FUNCTION_BLOCK "FB1062_HorDrillAutoStep"   // FB1062, SCL
{ S7_Optimized_Access := 'TRUE' }
// ============================================================
//  Block: FB1062_HorDrillAutoStep
//  ============================================================
//  编号：FB1062
//  原始语言：LAD（规则翻译为 SCL）
//  含义：Added Visual Chiseling Modeby WXY, 20220727
   VAR
      Aux : Struct   // 静态变量
         StartDrill : Bool;   // 静态变量
         DrillDepthMid : DInt;   // 打孔深度中间变量
         DrillDepthMax : Real;   // 静态变量
         DrillDepthMin : Real;   // 静态变量
         ScrLen_Mid : DInt;   // 批头长度中间变量
         OffSetYMid : DInt;   // 静态变量
         OffSetZMid : DInt;   // 静态变量
         go_X : Real;   // 机器人当前X位置
         go_Z : Real;   // 机器人当前Z位置
         MidPos_X : DInt;   // 静态变量
         MidPos_Z : DInt;   // 静态变量
         RobotSpeed : DInt;   // 机器人速度写入
         PressureMid : Real;   // 力中间变量
         HDrillOutTime : IEC_TIMER;   // 水平钻孔超时
         HStartTime : IEC_TIMER;   // 水平钻孔超时
      END_STRUCT;
      EdgeDetc : Struct   // 静态变量
         Pulse : Array[0..15] of Bool;   // 静态变量
      END_STRUCT;
      HorDrillStep : Struct   // 水平钻孔
         Busy : Bool;   // 静态变量
         StartCmd : Bool;   // 静态变量
         OKToStart : Bool;   // 静态变量
         TaskDone : Bool;   // 静态变量
         StepStart : Bool;   // 静态变量
         StepEnd : Bool;   // 静态变量
         ErrEnd : Bool;   // 静态变量
         ByPass : Bool;   // 静态变量
         TaskIO : Bool;   // 静态变量
         TaskNIO : Bool;   // 静态变量
         S1 : Bool;   // 静态变量
         S2 : Bool;   // 静态变量
         S3 : Bool;   // 静态变量
         S4 : Bool;   // 静态变量
         S5 : Bool;   // 静态变量
         S6 : Bool;   // 静态变量
         S7 : Bool;   // 静态变量
         S8 : Bool;   // 静态变量
         S9 : Bool;   // 静态变量
         S10 : Bool;   // 静态变量
         S11 : Bool;   // 静态变量
         S12 : Bool;   // 静态变量
         S13 : Bool;   // 静态变量
         S14 : Bool;   // 静态变量
         S15 : Bool;   // 静态变量
         S16 : Bool;   // 静态变量
         S17 : Bool;   // 静态变量
         S18 : Bool;   // 静态变量
         S19 : Bool;   // 静态变量
         S20 : Bool;   // 静态变量
         S21 : Bool;   // 静态变量
         S22 : Bool;   // 静态变量
         S23 : Bool;   // 静态变量
         S24 : Bool;   // 静态变量
         S25 : Bool;   // 静态变量
         S26 : Bool;   // 静态变量
         S27 : Bool;   // 静态变量
         S28 : Bool;   // 静态变量
         S29 : Bool;   // 静态变量
         S30 : Bool;   // 静态变量
         S31 : Bool;   // 静态变量
         S32 : Bool;   // 静态变量
         S33 : Bool;   // 静态变量
         S34 : Bool;   // 静态变量
         S35 : Bool;   // 静态变量
         S36 : Bool;   // 静态变量
         S37 : Bool;   // 静态变量
         S38 : Bool;   // 静态变量
         S39 : Bool;   // 静态变量
         S40 : Bool;   // 静态变量
         S41 : Bool;   // 静态变量
         S42 : Bool;   // 静态变量
         S43 : Bool;   // 静态变量
         S44 : Bool;   // 静态变量
         S45 : Bool;   // 静态变量
         S46 : Bool;   // 静态变量
         S47 : Bool;   // 静态变量
         S48 : Bool;   // 静态变量
         S49 : Bool;   // 静态变量
         S50 : Bool;   // 静态变量
         S51 : Bool;   // 静态变量
         S52 : Bool;   // 静态变量
         S53 : Bool;   // 静态变量
         S54 : Bool;   // 静态变量
         S55 : Bool;   // 静态变量
         S56 : Bool;   // 静态变量
         S57 : Bool;   // 静态变量
         S58 : Bool;   // 静态变量
         S59 : Bool;   // 静态变量
         S60 : Bool;   // 静态变量
         S61 : Bool;   // 静态变量
         S62 : Bool;   // 静态变量
         S63 : Bool;   // 静态变量
         S64 : Bool;   // 静态变量
         S65 : Bool;   // 静态变量
         S66 : Bool;   // 静态变量
         S67 : Bool;   // 静态变量
         StopDrill_Ack : Bool;   // 静态变量
         GougeStopDrill_Ack : Bool;   // 斜打结束请求
         StopDrill_End : Bool;   // 静态变量
         GougeStopDrill_End : Bool;   // 斜打异常结束请求
         InitForcePulse : Bool;   // 静态变量
      END_STRUCT;
      VisualOffsetMid : Struct   // 静态变量
         X : DInt;   // 静态变量
         Y : DInt;   // 静态变量
         Z : DInt;   // 静态变量
         "A" : DInt;   // 静态变量
         "B" : DInt;   // 静态变量
         C : DInt;   // 静态变量
         A0 : Real;   // 静态变量
         B0 : Real;   // 静态变量
         C0 : Real;   // 静态变量
      END_STRUCT;
      PT : Time;   // 静态变量
      ET : Time;   // 静态变量
      IN : Bool;   // 静态变量
      Q : Bool;   // 水平钻孔超时
   END_VAR
   VAR_TEMP
      StepPls : Bool;   // 临时变量
      HorPosMod : Int;   // 临时变量
   END_VAR
BEGIN

   // ---------- 网络 1 ----------
   // 标题：本工位必须要做(可能条件暂时不满足)
   // 含义：将 (("DB720_KuKa_MainCtrl".Ctrl_Out.RobotAction = 0) AND "DB720_KuKa_MainCtrl".Aux.ToolAtPos) AND NOT ("DB1148_PromptBeeper".Public.RobotNotReady) 赋给 #HorDrillStep.OKToStart
   #HorDrillStep.OKToStart := (("DB720_KuKa_MainCtrl".Ctrl_Out.RobotAction = 0) AND "DB720_KuKa_MainCtrl".Aux.ToolAtPos) AND NOT ("DB1148_PromptBeeper".Public.RobotNotReady);
   // 含义：条件 (("ManMode_M" AND "DB1900_Communication_PC".Recv.RobotDrillTPPB) AND ("DB1900_Communication_PC".Recv.ChooseProgNo = 1)) 成立时，将 TRUE 传送到 #HorDrillStep.StartCmd
   IF (("ManMode_M" AND "DB1900_Communication_PC".Recv.RobotDrillTPPB) AND ("DB1900_Communication_PC".Recv.ChooseProgNo = 1)) THEN
       #HorDrillStep.StartCmd := TRUE;
   END_IF;
   // 含义：将 "DB1900_Communication_PC".Para.DrillDepth; (* Convert → DInt *) END_IF 赋给 IF "DB1060_AutoStep".DownDrillAutoStep.DownDrillStep.StepStart THEN #Aux.DrillDepthMid
   IF "DB1060_AutoStep".DownDrillAutoStep.DownDrillStep.StepStart THEN
       #Aux.DrillDepthMid := "DB1900_Communication_PC".Para.DrillDepth; (* Convert → DInt *)
   END_IF;
   // 含义：将 SWAP(#Aux.DrillDepthMid) 赋给 "DB720_KuKa_MainCtrl".CmdOut.gi_Depth
   "DB720_KuKa_MainCtrl".CmdOut.gi_Depth := SWAP(#Aux.DrillDepthMid);
   // 含义：条件 #HorDrillStep.StepStart AND "DB1900_Communication_PC".Para.ProduceMode3 成立时，将 ("DB1900_Communication_PC".Para.DrillDepth + 0.0) 传送到 #Aux.DrillDepthMid
   IF #HorDrillStep.StepStart AND "DB1900_Communication_PC".Para.ProduceMode3 THEN
       #Aux.DrillDepthMid := ("DB1900_Communication_PC".Para.DrillDepth + 0.0);
   END_IF;
   // 含义：将 SWAP(#Aux.DrillDepthMid) 赋给 "DB720_KuKa_MainCtrl".CmdOut.gi_Depth
   "DB720_KuKa_MainCtrl".CmdOut.gi_Depth := SWAP(#Aux.DrillDepthMid);
   // 含义：条件 #HorDrillStep.StepStart AND "DB1900_Communication_PC".Para.ProduceMode3 成立时，将 "DB1910_DrillData".AUX.LayerNo 传送到 "DB720_KuKa_MainCtrl".CmdOut.gi_LayerNum
   IF #HorDrillStep.StepStart AND "DB1900_Communication_PC".Para.ProduceMode3 THEN
       "DB720_KuKa_MainCtrl".CmdOut.gi_LayerNum := "DB1910_DrillData".AUX.LayerNo;
   END_IF;
   // 含义：条件 #HorDrillStep.StepStart AND NOT ("DB1900_Communication_PC".Para.ProduceMode3) 成立时，将 ("DB1900_Communication_PC".Para.DrillDepth + 5.0) 传送到 #Aux.DrillDepthMid
   IF #HorDrillStep.StepStart AND NOT ("DB1900_Communication_PC".Para.ProduceMode3) THEN
       #Aux.DrillDepthMid := ("DB1900_Communication_PC".Para.DrillDepth + 5.0);
   END_IF;
   // 含义：将 SWAP(#Aux.DrillDepthMid) 赋给 "DB720_KuKa_MainCtrl".CmdOut.gi_Depth
   "DB720_KuKa_MainCtrl".CmdOut.gi_Depth := SWAP(#Aux.DrillDepthMid);
   // 含义：将 "DB1900_Communication_PC".Para.ScrLen; (* Convert → DInt *) 赋给 #Aux.ScrLen_Mid
   #Aux.ScrLen_Mid := "DB1900_Communication_PC".Para.ScrLen; (* Convert → DInt *)
   // 含义：将 SWAP(#Aux.ScrLen_Mid) 赋给 "DB720_KuKa_MainCtrl".CmdOut.gi_ScrewLength
   "DB720_KuKa_MainCtrl".CmdOut.gi_ScrewLength := SWAP(#Aux.ScrLen_Mid);

   // ---------- 网络 2 ----------
   // 标题：****************************机器人坐标数据传递 深度计算*********************************
   // 注释：Added Visual Chiseling Modeby WXY, 20220727
   // 含义：将 SWAP("DB720_KuKa_MainCtrl".StatusIn.go_X) 赋给 #Aux.MidPos_X
   #Aux.MidPos_X := SWAP("DB720_KuKa_MainCtrl".StatusIn.go_X);
   // 含义：将 #Aux.MidPos_X; (* Convert → Real *) 赋给 #Aux.go_X
   #Aux.go_X := #Aux.MidPos_X; (* Convert → Real *)
   // 含义：将 (#Aux.go_X / 1000.0) 赋给 "DB720_KuKa_MainCtrl".Aux.go_X
   "DB720_KuKa_MainCtrl".Aux.go_X := (#Aux.go_X / 1000.0);
   // 含义：将 SWAP("DB720_KuKa_MainCtrl".StatusIn.go_Z) 赋给 #Aux.MidPos_Z
   #Aux.MidPos_Z := SWAP("DB720_KuKa_MainCtrl".StatusIn.go_Z);
   // 含义：将 #Aux.MidPos_Z; (* Convert → Real *) 赋给 #Aux.go_Z
   #Aux.go_Z := #Aux.MidPos_Z; (* Convert → Real *)
   // 含义：将 (#Aux.go_Z / 1000.0) 赋给 "DB720_KuKa_MainCtrl".Aux.go_Z
   "DB720_KuKa_MainCtrl".Aux.go_Z := (#Aux.go_Z / 1000.0);
   // 含义：条件 (((#HorDrillStep.S12 AND "DB720_KuKa_MainCtrl".StatusIn.do_DrillReady_Act) AND "DB720_KuKa_MainCtrl".StatusIn.do_HorDril_Pos) OR (((((#HorDrillStep.S12 AND "DB720_KuKa_MainCtrl".StatusIn.do_DrillReady_Act) AND "DB2500 Visual Chiseling".VisualChiselingMode) AND "DB720_KuKa_MainCtrl".StatusIn.do_Gouge_Pos) AND ("DB1900_Communication_PC".Recv.Current_2 > "DB1900_Communication_PC".Para.CurrentMinLimit))) OR ((#HorDrillStep.S12 AND NOT (#HorDrillStep.S22)) AND #Aux.StartDrill)) AND NOT (#Aux.StartDrill) 成立时，将 "DB720_KuKa_MainCtrl".Aux.go_X 传送到 "DB720_KuKa_MainCtrl".Aux.XZeroPos
   IF (((#HorDrillStep.S12 AND "DB720_KuKa_MainCtrl".StatusIn.do_DrillReady_Act) AND "DB720_KuKa_MainCtrl".StatusIn.do_HorDril_Pos) OR (((((#HorDrillStep.S12 AND "DB720_KuKa_MainCtrl".StatusIn.do_DrillReady_Act) AND "DB2500 Visual Chiseling".VisualChiselingMode) AND "DB720_KuKa_MainCtrl".StatusIn.do_Gouge_Pos) AND ("DB1900_Communication_PC".Recv.Current_2 > "DB1900_Communication_PC".Para.CurrentMinLimit))) OR ((#HorDrillStep.S12 AND NOT (#HorDrillStep.S22)) AND #Aux.StartDrill)) AND NOT (#Aux.StartDrill) THEN
       "DB720_KuKa_MainCtrl".Aux.XZeroPos := "DB720_KuKa_MainCtrl".Aux.go_X;
   END_IF;
   // 含义：条件 ((#HorDrillStep.S12 AND "DB720_KuKa_MainCtrl".StatusIn.do_DrillReady_Act) AND "DB720_KuKa_MainCtrl".StatusIn.do_HorDril_Pos) OR (((((#HorDrillStep.S12 AND "DB720_KuKa_MainCtrl".StatusIn.do_DrillReady_Act) AND "DB2500 Visual Chiseling".VisualChiselingMode) AND "DB720_KuKa_MainCtrl".StatusIn.do_Gouge_Pos) AND ("DB1900_Communication_PC".Recv.Current_2 > "DB1900_Communication_PC".Para.CurrentMinLimit))) OR ((#HorDrillStep.S12 AND NOT (#HorDrillStep.S22)) AND #Aux.StartDrill) 成立时，将 ("DB720_KuKa_MainCtrl".Aux.go_X - "DB720_KuKa_MainCtrl".Aux.XZeroPos) 传送到 "DB720_KuKa_MainCtrl".Aux.CurrentRobPos
   IF ((#HorDrillStep.S12 AND "DB720_KuKa_MainCtrl".StatusIn.do_DrillReady_Act) AND "DB720_KuKa_MainCtrl".StatusIn.do_HorDril_Pos) OR (((((#HorDrillStep.S12 AND "DB720_KuKa_MainCtrl".StatusIn.do_DrillReady_Act) AND "DB2500 Visual Chiseling".VisualChiselingMode) AND "DB720_KuKa_MainCtrl".StatusIn.do_Gouge_Pos) AND ("DB1900_Communication_PC".Recv.Current_2 > "DB1900_Communication_PC".Para.CurrentMinLimit))) OR ((#HorDrillStep.S12 AND NOT (#HorDrillStep.S22)) AND #Aux.StartDrill) THEN
       "DB720_KuKa_MainCtrl".Aux.CurrentRobPos := ("DB720_KuKa_MainCtrl".Aux.go_X - "DB720_KuKa_MainCtrl".Aux.XZeroPos);
   END_IF;
   // 含义：将 ("DB720_KuKa_MainCtrl".Aux.CurrentRobPos - "DB1080_Component".ClinyderPos.Ctrl_Out.Cur_Val_Out) 赋给 "DB720_KuKa_MainCtrl".Aux.ScrLen_Mid1
   "DB720_KuKa_MainCtrl".Aux.ScrLen_Mid1 := ("DB720_KuKa_MainCtrl".Aux.CurrentRobPos - "DB1080_Component".ClinyderPos.Ctrl_Out.Cur_Val_Out);
   // 含义：条件 (("DB720_KuKa_MainCtrl".Aux.go_X >= "DB720_KuKa_MainCtrl".Aux.XZeroPos) AND ("DB720_KuKa_MainCtrl".Aux.ScrLen_Mid1 >= 0.0)) 成立时，将 "DB720_KuKa_MainCtrl".Aux.ScrLen_Mid1 传送到 "DB1900_Communication_PC".Send.ScrLen
   IF (("DB720_KuKa_MainCtrl".Aux.go_X >= "DB720_KuKa_MainCtrl".Aux.XZeroPos) AND ("DB720_KuKa_MainCtrl".Aux.ScrLen_Mid1 >= 0.0)) THEN
       "DB1900_Communication_PC".Send.ScrLen := "DB720_KuKa_MainCtrl".Aux.ScrLen_Mid1;
   END_IF;
   // 含义：条件 (((("DB720_KuKa_MainCtrl".Aux.go_X >= "DB720_KuKa_MainCtrl".Aux.XZeroPos) AND ("DB720_KuKa_MainCtrl".Aux.ScrLen_Mid1 <= 0.0))) AND ("DB1080_Component".ClinyderPos.Ctrl_Out.Cur_Val_Out >= 0.0)) 成立时，将 ABS("DB720_KuKa_MainCtrl".Aux.ScrLen_Mid1) 传送到 "DB1900_Communication_PC".Send.ScrLen
   IF (((("DB720_KuKa_MainCtrl".Aux.go_X >= "DB720_KuKa_MainCtrl".Aux.XZeroPos) AND ("DB720_KuKa_MainCtrl".Aux.ScrLen_Mid1 <= 0.0))) AND ("DB1080_Component".ClinyderPos.Ctrl_Out.Cur_Val_Out >= 0.0)) THEN
       "DB1900_Communication_PC".Send.ScrLen := ABS("DB720_KuKa_MainCtrl".Aux.ScrLen_Mid1);
   END_IF;
   // 含义：将 ((#HorDrillStep.S12 AND "DB720_KuKa_MainCtrl".StatusIn.do_DrillReady_Act) AND "DB720_KuKa_MainCtrl".StatusIn.do_HorDril_Pos) OR (((((#HorDrillStep.S12 AND "DB720_KuKa_MainCtrl".StatusIn.do_DrillReady_Act) AND "DB2500 Visual Chiseling".VisualChiselingMode) AND "DB720_KuKa_MainCtrl".StatusIn.do_Gouge_Pos) AND ("DB1900_Communication_PC".Recv.Current_2 > "DB1900_Communication_PC".Para.CurrentMinLimit))) OR ((#HorDrillStep.S12 AND NOT (#HorDrillStep.S22)) AND #Aux.StartDrill) 赋给 #Aux.StartDrill
   #Aux.StartDrill := ((#HorDrillStep.S12 AND "DB720_KuKa_MainCtrl".StatusIn.do_DrillReady_Act) AND "DB720_KuKa_MainCtrl".StatusIn.do_HorDril_Pos) OR (((((#HorDrillStep.S12 AND "DB720_KuKa_MainCtrl".StatusIn.do_DrillReady_Act) AND "DB2500 Visual Chiseling".VisualChiselingMode) AND "DB720_KuKa_MainCtrl".StatusIn.do_Gouge_Pos) AND ("DB1900_Communication_PC".Recv.Current_2 > "DB1900_Communication_PC".Para.CurrentMinLimit))) OR ((#HorDrillStep.S12 AND NOT (#HorDrillStep.S22)) AND #Aux.StartDrill);
   // 含义：调用计数器实例 "DB1042_Timer".HDrillEndTime.TON（上升沿计数，当前值写入 CV）
   "DB1042_Timer".HDrillEndTime.TON(IN := ((#HorDrillStep.S12 AND "DB720_KuKa_MainCtrl".StatusIn.do_DrillReady_Act) AND "DB720_KuKa_MainCtrl".StatusIn.do_HorDril_Pos) OR (((((#HorDrillStep.S12 AND "DB720_KuKa_MainCtrl".StatusIn.do_DrillReady_Act) AND "DB2500 Visual Chiseling".VisualChiselingMode) AND "DB720_KuKa_MainCtrl".StatusIn.do_Gouge_Pos) AND ("DB1900_Communication_PC".Recv.Current_2 > "DB1900_Communication_PC".Para.CurrentMinLimit))) OR ((#HorDrillStep.S12 AND NOT (#HorDrillStep.S22)) AND #Aux.StartDrill),
                                    PT := "DB1900_Communication_PC".Para.DrillTime);

   // ---------- 网络 3 ----------
   // 标题：************************************力计算*******************************************
   // 含义：条件 ("DB1900_Communication_PC".Send.ScrLen < 0.0) 成立时，将 0.0 传送到 "DB1900_Communication_PC".Send.ScrLen
   IF ("DB1900_Communication_PC".Send.ScrLen < 0.0) THEN
       "DB1900_Communication_PC".Send.ScrLen := 0.0;
   END_IF;
   // 含义：条件 ((("ManMode_M" AND NOT ("DB720_KuKa_MainCtrl".CheckBit.StepStart)) AND "DB2500 Visual Chiseling".RobotRetHomeCmd_AllMode) AND "DB1900_Communication_PC".Para.DrillDirection1) OR ((("ManMode_M" AND NOT ("DB720_KuKa_MainCtrl".CheckBit.StepStart)) AND "DB2500 Visual Chiseling".RobotRetHomeCmd_AllMode) AND "DB1900_Communication_PC".Para.DrillDirection2) 成立时，将 0.0 传送到 "DB1080_Component".Aux.Pressure
   IF ((("ManMode_M" AND NOT ("DB720_KuKa_MainCtrl".CheckBit.StepStart)) AND "DB2500 Visual Chiseling".RobotRetHomeCmd_AllMode) AND "DB1900_Communication_PC".Para.DrillDirection1) OR ((("ManMode_M" AND NOT ("DB720_KuKa_MainCtrl".CheckBit.StepStart)) AND "DB2500 Visual Chiseling".RobotRetHomeCmd_AllMode) AND "DB1900_Communication_PC".Para.DrillDirection2) THEN
       "DB1080_Component".Aux.Pressure := 0.0;
   END_IF;
   // 含义：条件 (("ManMode_M" AND NOT ("DB720_KuKa_MainCtrl".CheckBit.StepStart)) AND "DB2500 Visual Chiseling".RobotRetHomeCmd_AllMode) AND "DB1900_Communication_PC".Para.DrillDirection3 成立时，将 0.0 传送到 "DB1080_Component".Aux.Pressure
   IF (("ManMode_M" AND NOT ("DB720_KuKa_MainCtrl".CheckBit.StepStart)) AND "DB2500 Visual Chiseling".RobotRetHomeCmd_AllMode) AND "DB1900_Communication_PC".Para.DrillDirection3 THEN
       "DB1080_Component".Aux.Pressure := 0.0;
   END_IF;
   // 含义：条件 "ManMode_M" AND NOT ("DB720_KuKa_MainCtrl".CheckBit.StepStart) 成立时，将 FALSE 传送到 "DB720_KuKa_MainCtrl".CmdOut.di_ChiselCylinderRet
   IF "ManMode_M" AND NOT ("DB720_KuKa_MainCtrl".CheckBit.StepStart) THEN
       "DB720_KuKa_MainCtrl".CmdOut.di_ChiselCylinderRet := FALSE;
   END_IF;
   // 含义：条件 "ManMode_M" AND NOT ("DB720_KuKa_MainCtrl".CheckBit.StepStart) 成立时，将 FALSE 传送到 "DB720_KuKa_MainCtrl".CmdOut.di_ChiselRobotRet
   IF "ManMode_M" AND NOT ("DB720_KuKa_MainCtrl".CheckBit.StepStart) THEN
       "DB720_KuKa_MainCtrl".CmdOut.di_ChiselRobotRet := FALSE;
   END_IF;
   // 含义：条件 ("ManMode_M" AND NOT ("DB720_KuKa_MainCtrl".CheckBit.StepStart)) AND NOT ("DB2500 Visual Chiseling".RobotRetHomeCmd_AllMode) 成立时，将 0.3 传送到 "DB1080_Component".Aux.Pressure
   IF ("ManMode_M" AND NOT ("DB720_KuKa_MainCtrl".CheckBit.StepStart)) AND NOT ("DB2500 Visual Chiseling".RobotRetHomeCmd_AllMode) THEN
       "DB1080_Component".Aux.Pressure := 0.3;
   END_IF;

   // ---------- 网络 4 ----------
   // 标题：*********************************打孔超时及卡死计时*****************************************
   // 含义：调用定时器实例 #Aux.HDrillOutTime.TON
   #Aux.HDrillOutTime.TON(IN := "DB720_KuKa_MainCtrl".StatusIn.do_HorDril_Pos AND NOT ("DB1148_PromptBeeper".Public.DrillTimeOut),
                          PT := "DB1900_Communication_PC".Para.TimeOut);
   // 含义：调用定时器实例 "DB1042_Timer".GougeTimeOut.TON
   "DB1042_Timer".GougeTimeOut.TON(IN := ("DB720_KuKa_MainCtrl".StatusIn.do_Gouge_Pos OR "DB720_KuKa_MainCtrl".StatusIn.do_DrilEnd_Pos) AND NOT ("DB1148_PromptBeeper".Public.DrillTimeOut),
                                   PT := "DB1900_Communication_PC".Para.TimeOut);
   // 含义：调用计数器实例 "DB1042_Timer".CurrentLowTimeOut.TON（上升沿计数，当前值写入 CV）
   "DB1042_Timer".CurrentLowTimeOut.TON(IN := ((("DB720_KuKa_MainCtrl".StatusIn.do_HorDril_Pos OR "DB720_KuKa_MainCtrl".StatusIn.do_DownDril_Pos OR "DB720_KuKa_MainCtrl".StatusIn.do_JDiamond_MidPos OR "DB720_KuKa_MainCtrl".StatusIn.do_Gouge_Pos OR "DB720_KuKa_MainCtrl".StatusIn.do_DrilEnd_Pos) AND NOT ("DB1148_PromptBeeper".Public.DrillTimeOut)) AND ("DB1900_Communication_PC".Recv.Current_2 < "DB1900_Communication_PC".Para.CurrentMinLimit)),
                                        PT := "DB1900_Communication_PC".Para.CurrentMinLimitTimeOut);
   // 含义：调用计数器实例 "DB1042_Timer".CurrentHighTimeOut.TON（上升沿计数，当前值写入 CV）
   "DB1042_Timer".CurrentHighTimeOut.TON(IN := ((("DB720_KuKa_MainCtrl".StatusIn.do_HorDril_Pos OR "DB720_KuKa_MainCtrl".StatusIn.do_DownDril_Pos OR "DB720_KuKa_MainCtrl".StatusIn.do_JDiamond_MidPos OR "DB720_KuKa_MainCtrl".StatusIn.do_Gouge_Pos OR "DB720_KuKa_MainCtrl".StatusIn.do_DrilEnd_Pos) AND NOT ("DB1148_PromptBeeper".Public.DrillTimeOut)) AND ("DB1900_Communication_PC".Recv.Current_2 >= "DB1900_Communication_PC".Para.CurrentMaxLimit)),
                                         PT := T#200MS);
   // 含义：调用计数器实例 "DB1042_Timer".DrillingHighCurrentOut.TON（上升沿计数，当前值写入 CV）
   "DB1042_Timer".DrillingHighCurrentOut.TON(IN := (("DB720_KuKa_MainCtrl".StatusIn.do_HorDril_Pos OR "DB720_KuKa_MainCtrl".StatusIn.do_DownDril_Pos OR "DB720_KuKa_MainCtrl".StatusIn.do_JDiamond_MidPos OR "DB720_KuKa_MainCtrl".StatusIn.do_Gouge_Pos OR "DB720_KuKa_MainCtrl".StatusIn.do_DrilEnd_Pos) AND ("DB1900_Communication_PC".Recv.Current_2 >= "DB1900_Communication_PC".Para.CurrentMaxLimit)),
                                             PT := T#400MS);
   // 含义：调用定时器实例 "DB1042_Timer".FixtureStuckTimeOut.TON
   "DB1042_Timer".FixtureStuckTimeOut.TON(IN := ((((((("DB720_KuKa_MainCtrl".StatusIn.do_HorDril_Pos OR "DB720_KuKa_MainCtrl".StatusIn.do_DownDril_Pos OR "DB720_KuKa_MainCtrl".StatusIn.do_JDiamond_MidPos) AND NOT ("DB1900_Communication_PC".Para.ProduceMode3)) AND "AutoMode_M") OR (("DB1040_HomePos".MainStep.Start AND "IToolAtPos") AND "ManMode_M")) AND "DB1042_Timer".DrillMemory) AND NOT ("IFixtureStuckSensor")) AND ("DB720_KuKa_MainCtrl".CmdOut.gi_ToolTypeNo = 2)),
                                          PT := T#300MS);

   // ---------- 网络 5 ----------
   // 标题：**********************************钻孔区间*******************************************
   // 含义：将 ("DB1900_Communication_PC".Para.DrillDepth + 10.0) 赋给 #Aux.DrillDepthMax
   #Aux.DrillDepthMax := ("DB1900_Communication_PC".Para.DrillDepth + 10.0);
   // 含义：将 ("DB1900_Communication_PC".Para.DrillDepth - 5.0) 赋给 #Aux.DrillDepthMin
   #Aux.DrillDepthMin := ("DB1900_Communication_PC".Para.DrillDepth - 5.0);

   // ---------- 网络 6 ----------
   // 标题：*********************************水平钻孔Start****************************************
   // 含义：将 (((((((#HorDrillStep.StartCmd AND #HorDrillStep.OKToStart) OR #HorDrillStep.StepStart) AND "AllMode_M") AND "DB1900_Communication_PC".Recv.Z05ExtTPPB) AND ("DB1900_Communication_PC".Recv.Current_2 >= 0.5))) AND NOT ("DB1900_Communication_PC".Recv.EmmMode)) AND NOT (#HorDrillStep.StepEnd) 赋给 #HorDrillStep.StepStart
   #HorDrillStep.StepStart := (((((((#HorDrillStep.StartCmd AND #HorDrillStep.OKToStart) OR #HorDrillStep.StepStart) AND "AllMode_M") AND "DB1900_Communication_PC".Recv.Z05ExtTPPB) AND ("DB1900_Communication_PC".Recv.Current_2 >= 0.5))) AND NOT ("DB1900_Communication_PC".Recv.EmmMode)) AND NOT (#HorDrillStep.StepEnd);
   // 含义：将 (((((((#HorDrillStep.StartCmd AND #HorDrillStep.OKToStart) OR #HorDrillStep.StepStart) AND "AllMode_M") AND "DB1900_Communication_PC".Recv.Z05ExtTPPB) AND ("DB1900_Communication_PC".Recv.Current_2 >= 0.5))) AND NOT ("DB1900_Communication_PC".Recv.EmmMode)) AND NOT (#HorDrillStep.StepEnd) 赋给 #HorDrillStep.Busy
   #HorDrillStep.Busy := (((((((#HorDrillStep.StartCmd AND #HorDrillStep.OKToStart) OR #HorDrillStep.StepStart) AND "AllMode_M") AND "DB1900_Communication_PC".Recv.Z05ExtTPPB) AND ("DB1900_Communication_PC".Recv.Current_2 >= 0.5))) AND NOT ("DB1900_Communication_PC".Recv.EmmMode)) AND NOT (#HorDrillStep.StepEnd);
   // 含义：调用计数器实例 #Aux.HStartTime.TON（上升沿计数，当前值写入 CV）
   #Aux.HStartTime.TON(IN := (((((((#HorDrillStep.StartCmd AND #HorDrillStep.OKToStart) OR #HorDrillStep.StepStart) AND "AllMode_M") AND "DB1900_Communication_PC".Recv.Z05ExtTPPB) AND ("DB1900_Communication_PC".Recv.Current_2 >= 0.5))) AND NOT ("DB1900_Communication_PC".Recv.EmmMode)) AND NOT (#HorDrillStep.StepEnd),
                       PT := T#20S);
   // 含义：条件 NOT ((((((((#HorDrillStep.StartCmd AND #HorDrillStep.OKToStart) OR #HorDrillStep.StepStart) AND "AllMode_M") AND "DB1900_Communication_PC".Recv.Z05ExtTPPB) AND ("DB1900_Communication_PC".Recv.Current_2 >= 0.5))) AND NOT ("DB1900_Communication_PC".Recv.EmmMode)) AND NOT (#HorDrillStep.StepEnd)) 成立时，将 FALSE 传送到 #HorDrillStep.StopDrill_Ack
   IF NOT ((((((((#HorDrillStep.StartCmd AND #HorDrillStep.OKToStart) OR #HorDrillStep.StepStart) AND "AllMode_M") AND "DB1900_Communication_PC".Recv.Z05ExtTPPB) AND ("DB1900_Communication_PC".Recv.Current_2 >= 0.5))) AND NOT ("DB1900_Communication_PC".Recv.EmmMode)) AND NOT (#HorDrillStep.StepEnd)) THEN
       #HorDrillStep.StopDrill_Ack := FALSE;
   END_IF;
   // 含义：条件 NOT ((((((((#HorDrillStep.StartCmd AND #HorDrillStep.OKToStart) OR #HorDrillStep.StepStart) AND "AllMode_M") AND "DB1900_Communication_PC".Recv.Z05ExtTPPB) AND ("DB1900_Communication_PC".Recv.Current_2 >= 0.5))) AND NOT ("DB1900_Communication_PC".Recv.EmmMode)) AND NOT (#HorDrillStep.StepEnd)) 成立时，将 FALSE 传送到 #HorDrillStep.ErrEnd
   IF NOT ((((((((#HorDrillStep.StartCmd AND #HorDrillStep.OKToStart) OR #HorDrillStep.StepStart) AND "AllMode_M") AND "DB1900_Communication_PC".Recv.Z05ExtTPPB) AND ("DB1900_Communication_PC".Recv.Current_2 >= 0.5))) AND NOT ("DB1900_Communication_PC".Recv.EmmMode)) AND NOT (#HorDrillStep.StepEnd)) THEN
       #HorDrillStep.ErrEnd := FALSE;
   END_IF;

   // ---------- 网络 7 ----------
   // 标题：初始化
   // 注释：Added DB2700.VisualChiselingStart  by WXY, 20220615.
   // 含义：条件 (#HorDrillStep.StepStart AND NOT (#HorDrillStep.ErrEnd)) AND NOT (#HorDrillStep.S1) 成立时，将 FALSE 传送到 #HorDrillStep.TaskIO
   IF (#HorDrillStep.StepStart AND NOT (#HorDrillStep.ErrEnd)) AND NOT (#HorDrillStep.S1) THEN
       #HorDrillStep.TaskIO := FALSE;
   END_IF;
   // 含义：条件 (#HorDrillStep.StepStart AND NOT (#HorDrillStep.ErrEnd)) AND NOT (#HorDrillStep.S1) 成立时，将 FALSE 传送到 #HorDrillStep.TaskNIO
   IF (#HorDrillStep.StepStart AND NOT (#HorDrillStep.ErrEnd)) AND NOT (#HorDrillStep.S1) THEN
       #HorDrillStep.TaskNIO := FALSE;
   END_IF;
   // 含义：条件 (#HorDrillStep.StepStart AND NOT (#HorDrillStep.ErrEnd)) AND NOT (#HorDrillStep.S1) 成立时，将 FALSE 传送到 "DB720_KuKa_MainCtrl".CmdOut.di_ChiselCylinderRet
   IF (#HorDrillStep.StepStart AND NOT (#HorDrillStep.ErrEnd)) AND NOT (#HorDrillStep.S1) THEN
       "DB720_KuKa_MainCtrl".CmdOut.di_ChiselCylinderRet := FALSE;
   END_IF;
   // 含义：条件 (#HorDrillStep.StepStart AND NOT (#HorDrillStep.ErrEnd)) AND NOT (#HorDrillStep.S1) 成立时，将 FALSE 传送到 "DB720_KuKa_MainCtrl".CmdOut.di_ChiselRobotRet
   IF (#HorDrillStep.StepStart AND NOT (#HorDrillStep.ErrEnd)) AND NOT (#HorDrillStep.S1) THEN
       "DB720_KuKa_MainCtrl".CmdOut.di_ChiselRobotRet := FALSE;
   END_IF;
   // 含义：条件 (#HorDrillStep.StepStart AND NOT (#HorDrillStep.ErrEnd)) AND NOT (#HorDrillStep.S1) 成立时，将 FALSE 传送到 #HorDrillStep.StopDrill_Ack
   IF (#HorDrillStep.StepStart AND NOT (#HorDrillStep.ErrEnd)) AND NOT (#HorDrillStep.S1) THEN
       #HorDrillStep.StopDrill_Ack := FALSE;
   END_IF;
   // 含义：条件 (#HorDrillStep.StepStart AND NOT (#HorDrillStep.ErrEnd)) AND NOT (#HorDrillStep.S1) 成立时，将 1 传送到 "DB720_KuKa_MainCtrl".Aux.ForceNum
   IF (#HorDrillStep.StepStart AND NOT (#HorDrillStep.ErrEnd)) AND NOT (#HorDrillStep.S1) THEN
       "DB720_KuKa_MainCtrl".Aux.ForceNum := 1;
   END_IF;
   // 含义：将 #HorDrillStep.StepStart AND NOT (#HorDrillStep.ErrEnd) 赋给 #HorDrillStep.S1
   #HorDrillStep.S1 := #HorDrillStep.StepStart AND NOT (#HorDrillStep.ErrEnd);
   // 含义：条件 ((#HorDrillStep.StepStart AND NOT (#HorDrillStep.ErrEnd)) AND "DB2500 Visual Chiseling".VisualChiselingMode) AND "DB2500 Visual Chiseling".VisualCameraEnd 成立时，将 TRUE 传送到 "DB2500 Visual Chiseling".VisualChiselingStart
   IF ((#HorDrillStep.StepStart AND NOT (#HorDrillStep.ErrEnd)) AND "DB2500 Visual Chiseling".VisualChiselingMode) AND "DB2500 Visual Chiseling".VisualCameraEnd THEN
       "DB2500 Visual Chiseling".VisualChiselingStart := TRUE;
   END_IF;
   // 含义：条件 ((#HorDrillStep.StepStart AND NOT (#HorDrillStep.ErrEnd)) AND "DB2500 Visual Chiseling".VisualChiselingMode) AND "DB2500 Visual Chiseling".VisualCameraEnd 成立时，将 FALSE 传送到 "DB2500 Visual Chiseling".VisualChiselingEnd
   IF ((#HorDrillStep.StepStart AND NOT (#HorDrillStep.ErrEnd)) AND "DB2500 Visual Chiseling".VisualChiselingMode) AND "DB2500 Visual Chiseling".VisualCameraEnd THEN
       "DB2500 Visual Chiseling".VisualChiselingEnd := FALSE;
   END_IF;

   // ---------- 网络 8 ----------
   // 标题：判断条件
   // 含义：将 (#HorDrillStep.S1 AND NOT ("DB1147_PromptStartNotPmt".Public.ChangeHorDrillSlab)) OR (#HorDrillStep.S1 AND NOT ("DB1147_PromptStartNotPmt".Public.ChangeHorVChiselSlab)) OR (#HorDrillStep.S1 AND #HorDrillStep.S2) 赋给 #HorDrillStep.S2
   #HorDrillStep.S2 := (#HorDrillStep.S1 AND NOT ("DB1147_PromptStartNotPmt".Public.ChangeHorDrillSlab)) OR (#HorDrillStep.S1 AND NOT ("DB1147_PromptStartNotPmt".Public.ChangeHorVChiselSlab)) OR (#HorDrillStep.S1 AND #HorDrillStep.S2);
   // 含义：条件 ((#HorDrillStep.S1 AND "DB1147_PromptStartNotPmt".Public.ChangeHorDrillSlab) AND NOT ("DB2500 Visual Chiseling".VisualChiselingMode)) OR ((#HorDrillStep.S1 AND "DB1147_PromptStartNotPmt".Public.ChangeHorVChiselSlab) AND "DB2500 Visual Chiseling".VisualChiselingMode) 成立时，将 TRUE 传送到 #HorDrillStep.ErrEnd
   IF ((#HorDrillStep.S1 AND "DB1147_PromptStartNotPmt".Public.ChangeHorDrillSlab) AND NOT ("DB2500 Visual Chiseling".VisualChiselingMode)) OR ((#HorDrillStep.S1 AND "DB1147_PromptStartNotPmt".Public.ChangeHorVChiselSlab) AND "DB2500 Visual Chiseling".VisualChiselingMode) THEN
       #HorDrillStep.ErrEnd := TRUE;
   END_IF;

   // ---------- 网络 9 ----------
   // 标题：电源夹具ID号错误，请检查夹具！
   // 含义：将 ((((#HorDrillStep.S2 AND ("DB1900_Communication_PC".Para.IOFixtureNo = "DB1080_Component".IOFixtureIID.TP_CurFixtureID))) AND ("DB1900_Communication_PC".Para.PowerFixtureNo = "DB1080_Component".PowerFixtureID.TP_CurFixtureID))) OR (#HorDrillStep.S2 AND #HorDrillStep.S5) 赋给 #HorDrillStep.S5
   #HorDrillStep.S5 := ((((#HorDrillStep.S2 AND ("DB1900_Communication_PC".Para.IOFixtureNo = "DB1080_Component".IOFixtureIID.TP_CurFixtureID))) AND ("DB1900_Communication_PC".Para.PowerFixtureNo = "DB1080_Component".PowerFixtureID.TP_CurFixtureID))) OR (#HorDrillStep.S2 AND #HorDrillStep.S5);

   // ---------- 网络 10 ----------
   // 标题：推力气缸
   // 含义：条件 (#HorDrillStep.S5 AND NOT (#HorDrillStep.S7)) OR ((#HorDrillStep.S5 AND "DB2500 Visual Chiseling".VisualChiselingMode) AND "DB720_KuKa_MainCtrl".StatusIn.do_ChiselCylinderExt) 成立时，将 TRUE 传送到 "DB1081_ValveCall".ST01.Z01.ExtAuto
   IF (#HorDrillStep.S5 AND NOT (#HorDrillStep.S7)) OR ((#HorDrillStep.S5 AND "DB2500 Visual Chiseling".VisualChiselingMode) AND "DB720_KuKa_MainCtrl".StatusIn.do_ChiselCylinderExt) THEN
       "DB1081_ValveCall".ST01.Z01.ExtAuto := TRUE;
   END_IF;
   // 含义：条件 (#HorDrillStep.S5 AND NOT (#HorDrillStep.S7)) OR ((#HorDrillStep.S5 AND "DB2500 Visual Chiseling".VisualChiselingMode) AND "DB720_KuKa_MainCtrl".StatusIn.do_ChiselCylinderExt) 成立时，将 TRUE 传送到 "DB1081_ValveCall".ST01.Z02.VentValveAuto
   IF (#HorDrillStep.S5 AND NOT (#HorDrillStep.S7)) OR ((#HorDrillStep.S5 AND "DB2500 Visual Chiseling".VisualChiselingMode) AND "DB720_KuKa_MainCtrl".StatusIn.do_ChiselCylinderExt) THEN
       "DB1081_ValveCall".ST01.Z02.VentValveAuto := TRUE;
   END_IF;
   // 含义：条件 (#HorDrillStep.S5 AND NOT (#HorDrillStep.S7)) OR ((#HorDrillStep.S5 AND "DB2500 Visual Chiseling".VisualChiselingMode) AND "DB720_KuKa_MainCtrl".StatusIn.do_ChiselCylinderExt) 成立时，将 TRUE 传送到 "DB1081_ValveCall".ST01.Z05.ExtAuto
   IF (#HorDrillStep.S5 AND NOT (#HorDrillStep.S7)) OR ((#HorDrillStep.S5 AND "DB2500 Visual Chiseling".VisualChiselingMode) AND "DB720_KuKa_MainCtrl".StatusIn.do_ChiselCylinderExt) THEN
       "DB1081_ValveCall".ST01.Z05.ExtAuto := TRUE;
   END_IF;
   // 含义：条件 (#HorDrillStep.S5 AND NOT (#HorDrillStep.S7)) OR ((#HorDrillStep.S5 AND "DB2500 Visual Chiseling".VisualChiselingMode) AND "DB720_KuKa_MainCtrl".StatusIn.do_ChiselCylinderExt) 成立时，将 TRUE 传送到 "DB1081_ValveCall".ST01.Z06.RetAuto
   IF (#HorDrillStep.S5 AND NOT (#HorDrillStep.S7)) OR ((#HorDrillStep.S5 AND "DB2500 Visual Chiseling".VisualChiselingMode) AND "DB720_KuKa_MainCtrl".StatusIn.do_ChiselCylinderExt) THEN
       "DB1081_ValveCall".ST01.Z06.RetAuto := TRUE;
   END_IF;
   // 含义：条件 ((((#HorDrillStep.S5 AND NOT (#HorDrillStep.S7)) OR ((#HorDrillStep.S5 AND "DB2500 Visual Chiseling".VisualChiselingMode) AND "DB720_KuKa_MainCtrl".StatusIn.do_ChiselCylinderExt)) AND ("DB720_KuKa_MainCtrl".CmdOut.gi_ToolTypeNo = 13))) AND TRUE 成立时，将 TRUE 传送到 "QCamCoverExt"
   IF ((((#HorDrillStep.S5 AND NOT (#HorDrillStep.S7)) OR ((#HorDrillStep.S5 AND "DB2500 Visual Chiseling".VisualChiselingMode) AND "DB720_KuKa_MainCtrl".StatusIn.do_ChiselCylinderExt)) AND ("DB720_KuKa_MainCtrl".CmdOut.gi_ToolTypeNo = 13))) AND TRUE THEN
       "QCamCoverExt" := TRUE;
   END_IF;
   // 含义：条件 ((((#HorDrillStep.S5 AND NOT (#HorDrillStep.S7)) OR ((#HorDrillStep.S5 AND "DB2500 Visual Chiseling".VisualChiselingMode) AND "DB720_KuKa_MainCtrl".StatusIn.do_ChiselCylinderExt)) AND ("DB720_KuKa_MainCtrl".CmdOut.gi_ToolTypeNo = 13))) AND TRUE 成立时，将 FALSE 传送到 "QCamCoverRet"
   IF ((((#HorDrillStep.S5 AND NOT (#HorDrillStep.S7)) OR ((#HorDrillStep.S5 AND "DB2500 Visual Chiseling".VisualChiselingMode) AND "DB720_KuKa_MainCtrl".StatusIn.do_ChiselCylinderExt)) AND ("DB720_KuKa_MainCtrl".CmdOut.gi_ToolTypeNo = 13))) AND TRUE THEN
       "QCamCoverRet" := FALSE;
   END_IF;
   // 含义：条件 (#HorDrillStep.S5 AND NOT (#HorDrillStep.S7)) OR ((#HorDrillStep.S5 AND "DB2500 Visual Chiseling".VisualChiselingMode) AND "DB720_KuKa_MainCtrl".StatusIn.do_ChiselCylinderExt) 成立时，将 0.0 传送到 "DB1900_Communication_PC".Send.ScrLen
   IF (#HorDrillStep.S5 AND NOT (#HorDrillStep.S7)) OR ((#HorDrillStep.S5 AND "DB2500 Visual Chiseling".VisualChiselingMode) AND "DB720_KuKa_MainCtrl".StatusIn.do_ChiselCylinderExt) THEN
       "DB1900_Communication_PC".Send.ScrLen := 0.0;
   END_IF;
   // 含义：条件 (#HorDrillStep.S5 AND NOT (#HorDrillStep.S7)) OR ((#HorDrillStep.S5 AND "DB2500 Visual Chiseling".VisualChiselingMode) AND "DB720_KuKa_MainCtrl".StatusIn.do_ChiselCylinderExt) 成立时，将 0.3 传送到 "DB1080_Component".Aux.Pressure
   IF (#HorDrillStep.S5 AND NOT (#HorDrillStep.S7)) OR ((#HorDrillStep.S5 AND "DB2500 Visual Chiseling".VisualChiselingMode) AND "DB720_KuKa_MainCtrl".StatusIn.do_ChiselCylinderExt) THEN
       "DB1080_Component".Aux.Pressure := 0.3;
   END_IF;
   // 含义：条件 (#HorDrillStep.S5 AND "DB720_KuKa_MainCtrl".StatusIn.do_ReqDrilling) AND NOT ("DB2500 Visual Chiseling".VisualChiselingMode) 成立时，将 ( "DB1900_Communication_PC".Para.InitialForce + -55.1) / 1308.0 传送到 "DB1080_Component".Aux.Pressure
   IF (#HorDrillStep.S5 AND "DB720_KuKa_MainCtrl".StatusIn.do_ReqDrilling) AND NOT ("DB2500 Visual Chiseling".VisualChiselingMode) THEN
       "DB1080_Component".Aux.Pressure := ("DB1900_Communication_PC".Para.InitialForce + -55.1) / 1308.0;
   END_IF;
   // 含义：条件 (#HorDrillStep.S5 AND "DB720_KuKa_MainCtrl".StatusIn.do_ReqDrilling) AND "DB2500 Visual Chiseling".VisualChiselingMode 成立时，将 (30.0 + ("DB2500 Visual Chiseling".OffsetB_GravityComp)) 传送到 #Aux.PressureMid
   IF (#HorDrillStep.S5 AND "DB720_KuKa_MainCtrl".StatusIn.do_ReqDrilling) AND "DB2500 Visual Chiseling".VisualChiselingMode THEN
       #Aux.PressureMid := (30.0 + ("DB2500 Visual Chiseling".OffsetB_GravityComp));
   END_IF;
   // 含义：将 ( #Aux.PressureMid + -55.1) / 1308.0 赋给 "DB1080_Component".Aux.Pressure
   "DB1080_Component".Aux.Pressure := (#Aux.PressureMid + -55.1) / 1308.0;
   // 含义：将 ((((#HorDrillStep.S5 AND "DB1081_ValveCall".ST01.Z01.ExtPos) OR ((#HorDrillStep.S5 AND "DB1900_Communication_PC".Para.DrillDirection1) AND "DB1900_Communication_PC".Para.ProduceMode3)) AND "IZ02ExtPos") AND "DB1081_ValveCall".ST01.Z06.RetPos) OR (#HorDrillStep.S5 AND #HorDrillStep.S7) 赋给 #HorDrillStep.S7
   #HorDrillStep.S7 := ((((#HorDrillStep.S5 AND "DB1081_ValveCall".ST01.Z01.ExtPos) OR ((#HorDrillStep.S5 AND "DB1900_Communication_PC".Para.DrillDirection1) AND "DB1900_Communication_PC".Para.ProduceMode3)) AND "IZ02ExtPos") AND "DB1081_ValveCall".ST01.Z06.RetPos) OR (#HorDrillStep.S5 AND #HorDrillStep.S7);

   // ---------- 网络 11 ----------
   // 标题：数据写入 X宽 Y长  NOT Visual Chiseling Mode
   // 注释：Added Not Visual Chiseling Mode DB2500.DBX30.0 by WXY, 20220726. PosNo is ToolNo, not HoleNo.
   // 含义：将 "DB1910_DrillData".HorDrill.gi_OffSetY; (* Convert → DInt *) END_IF 赋给 IF (#HorDrillStep.S7 AND NOT ("DB2500 Visual Chiseling".VisualChiselingMode)) AND NOT (#HorDrillStep.S10) THEN #Aux.OffSetYMid
   IF (#HorDrillStep.S7 AND NOT ("DB2500 Visual Chiseling".VisualChiselingMode)) AND NOT (#HorDrillStep.S10) THEN
       #Aux.OffSetYMid := "DB1910_DrillData".HorDrill.gi_OffSetY; (* Convert → DInt *)
   END_IF;
   // 含义：将 SWAP(#Aux.OffSetYMid) 赋给 "DB720_KuKa_MainCtrl".CmdOut.gi_OffSetY
   "DB720_KuKa_MainCtrl".CmdOut.gi_OffSetY := SWAP(#Aux.OffSetYMid);
   // 含义：将 "DB1910_DrillData".HorDrill.gi_OffSetZ; (* Convert → DInt *) END_IF 赋给 IF (#HorDrillStep.S7 AND NOT ("DB2500 Visual Chiseling".VisualChiselingMode)) AND NOT (#HorDrillStep.S10) THEN #Aux.OffSetZMid
   IF (#HorDrillStep.S7 AND NOT ("DB2500 Visual Chiseling".VisualChiselingMode)) AND NOT (#HorDrillStep.S10) THEN
       #Aux.OffSetZMid := "DB1910_DrillData".HorDrill.gi_OffSetZ; (* Convert → DInt *)
   END_IF;
   // 含义：将 SWAP(#Aux.OffSetZMid) 赋给 "DB720_KuKa_MainCtrl".CmdOut.gi_OffSetZ
   "DB720_KuKa_MainCtrl".CmdOut.gi_OffSetZ := SWAP(#Aux.OffSetZMid);
   // 含义：将 #HorDrillStep.S7 AND NOT ("DB2500 Visual Chiseling".VisualChiselingMode) 赋给 #HorDrillStep.S10
   #HorDrillStep.S10 := #HorDrillStep.S7 AND NOT ("DB2500 Visual Chiseling".VisualChiselingMode);

   // ---------- 网络 12 ----------
   // 标题：辅助气缸
   // 注释：Added Visual Chiseling Mode DB2500.DBX30.0 by WXY, 20220726.   ( Always Send Offset Value in Visual Chiseling Mode)
   // 含义：将 (((((#HorDrillStep.S7 AND "DB2500 Visual Chiseling".VisualChiselingMode) OR #HorDrillStep.S10) AND "IZ02ExtPos") AND ("DB1080_Component".ClinyderPos.Ctrl_Out.Cur_Val_Out <= 1.0))) OR ((((#HorDrillStep.S7 AND "DB2500 Visual Chiseling".VisualChiselingMode) OR #HorDrillStep.S10) AND "DB1900_Communication_PC".Para.DrillDirection1) AND "DB1900_Communication_PC".Para.ProduceMode3) OR (((#HorDrillStep.S7 AND "DB2500 Visual Chiseling".VisualChiselingMode) OR #HorDrillStep.S10) AND #HorDrillStep.S12) 赋给 #HorDrillStep.S12
   #HorDrillStep.S12 := (((((#HorDrillStep.S7 AND "DB2500 Visual Chiseling".VisualChiselingMode) OR #HorDrillStep.S10) AND "IZ02ExtPos") AND ("DB1080_Component".ClinyderPos.Ctrl_Out.Cur_Val_Out <= 1.0))) OR ((((#HorDrillStep.S7 AND "DB2500 Visual Chiseling".VisualChiselingMode) OR #HorDrillStep.S10) AND "DB1900_Communication_PC".Para.DrillDirection1) AND "DB1900_Communication_PC".Para.ProduceMode3) OR (((#HorDrillStep.S7 AND "DB2500 Visual Chiseling".VisualChiselingMode) OR #HorDrillStep.S10) AND #HorDrillStep.S12);
   // 含义：条件 (((((((#HorDrillStep.S7 AND "DB2500 Visual Chiseling".VisualChiselingMode) OR #HorDrillStep.S10) AND "DB1900_Communication_PC".Para.DrillDirection1) AND "DB2500 Visual Chiseling".VisualChiselingMode) AND "IZ02ExtPos") AND "DB1081_ValveCall".ST01.Z01.ExtPos) AND ("DB1080_Component".ClinyderPos.Ctrl_Out.Cur_Val_Out <= 2.0)) 成立时，将 TRUE 传送到 "DB720_KuKa_MainCtrl".CmdOut.di_PushCylOK_Sig
   IF (((((((#HorDrillStep.S7 AND "DB2500 Visual Chiseling".VisualChiselingMode) OR #HorDrillStep.S10) AND "DB1900_Communication_PC".Para.DrillDirection1) AND "DB2500 Visual Chiseling".VisualChiselingMode) AND "IZ02ExtPos") AND "DB1081_ValveCall".ST01.Z01.ExtPos) AND ("DB1080_Component".ClinyderPos.Ctrl_Out.Cur_Val_Out <= 2.0)) THEN
       "DB720_KuKa_MainCtrl".CmdOut.di_PushCylOK_Sig := TRUE;
   END_IF;
   // 含义：条件 (((((#HorDrillStep.S7 AND "DB2500 Visual Chiseling".VisualChiselingMode) OR #HorDrillStep.S10) AND "DB1900_Communication_PC".Para.DrillDirection1) AND "DB2500 Visual Chiseling".VisualChiselingMode) AND ("DB1080_Component".ClinyderPos.Ctrl_Out.Cur_Val_Out > 2.0)) 成立时，将 FALSE 传送到 "DB720_KuKa_MainCtrl".CmdOut.di_PushCylOK_Sig
   IF (((((#HorDrillStep.S7 AND "DB2500 Visual Chiseling".VisualChiselingMode) OR #HorDrillStep.S10) AND "DB1900_Communication_PC".Para.DrillDirection1) AND "DB2500 Visual Chiseling".VisualChiselingMode) AND ("DB1080_Component".ClinyderPos.Ctrl_Out.Cur_Val_Out > 2.0)) THEN
       "DB720_KuKa_MainCtrl".CmdOut.di_PushCylOK_Sig := FALSE;
   END_IF;

   // ---------- 网络 13 ----------
   // 标题：调用机器人
   // 注释：Send ProgNo 15 to Robot in Visual Chiseling Mode by WXY, 20220615.
   // 含义：条件 (#HorDrillStep.S12 AND NOT (#HorDrillStep.S15)) AND "DB1900_Communication_PC".Para.ProduceMode2 成立时，将 1 传送到 "DB1080_Component".Robot.CTRL_IN.ProgNo
   IF (#HorDrillStep.S12 AND NOT (#HorDrillStep.S15)) AND "DB1900_Communication_PC".Para.ProduceMode2 THEN
       "DB1080_Component".Robot.CTRL_IN.ProgNo := 1;
   END_IF;
   // 含义：条件 (((#HorDrillStep.S12 AND NOT (#HorDrillStep.S15)) AND "DB1900_Communication_PC".Para.ProduceMode3) AND NOT ("DB2500 Visual Chiseling".VisualChiselingMode)) AND NOT ("DB1900_Communication_PC".Para.SwingOn) 成立时，将 13 传送到 "DB1080_Component".Robot.CTRL_IN.ProgNo
   IF (((#HorDrillStep.S12 AND NOT (#HorDrillStep.S15)) AND "DB1900_Communication_PC".Para.ProduceMode3) AND NOT ("DB2500 Visual Chiseling".VisualChiselingMode)) AND NOT ("DB1900_Communication_PC".Para.SwingOn) THEN
       "DB1080_Component".Robot.CTRL_IN.ProgNo := 13;
   END_IF;
   // 含义：条件 (((#HorDrillStep.S12 AND NOT (#HorDrillStep.S15)) AND "DB1900_Communication_PC".Para.ProduceMode3) AND NOT ("DB2500 Visual Chiseling".VisualChiselingMode)) AND "DB1900_Communication_PC".Para.SwingOn 成立时，将 14 传送到 "DB1080_Component".Robot.CTRL_IN.ProgNo
   IF (((#HorDrillStep.S12 AND NOT (#HorDrillStep.S15)) AND "DB1900_Communication_PC".Para.ProduceMode3) AND NOT ("DB2500 Visual Chiseling".VisualChiselingMode)) AND "DB1900_Communication_PC".Para.SwingOn THEN
       "DB1080_Component".Robot.CTRL_IN.ProgNo := 14;
   END_IF;
   // 含义：条件 ((#HorDrillStep.S12 AND NOT (#HorDrillStep.S15)) AND "DB1900_Communication_PC".Para.ProduceMode3) AND "DB2500 Visual Chiseling".VisualChiselingMode 成立时，将 15 传送到 "DB1080_Component".Robot.CTRL_IN.ProgNo
   IF ((#HorDrillStep.S12 AND NOT (#HorDrillStep.S15)) AND "DB1900_Communication_PC".Para.ProduceMode3) AND "DB2500 Visual Chiseling".VisualChiselingMode THEN
       "DB1080_Component".Robot.CTRL_IN.ProgNo := 15;
   END_IF;
   // 含义：条件 #HorDrillStep.S12 AND NOT (#HorDrillStep.S15) 成立时，将 50 传送到 "DB1080_Component".Robot.CTRL_IN.RobotSpeed
   IF #HorDrillStep.S12 AND NOT (#HorDrillStep.S15) THEN
       "DB1080_Component".Robot.CTRL_IN.RobotSpeed := 50;
   END_IF;
   // 含义：将 #HorDrillStep.S12 AND NOT (#HorDrillStep.S15) 赋给 "DB1146_PromptFree".Public.do_HorDril_Pos
   "DB1146_PromptFree".Public.do_HorDril_Pos := #HorDrillStep.S12 AND NOT (#HorDrillStep.S15);
   // 含义：条件 #HorDrillStep.S12 成立时，将 TRUE 传送到 "DB1080_Component".Robot.Cmd.Auto.ProgStart
   IF #HorDrillStep.S12 THEN
       "DB1080_Component".Robot.Cmd.Auto.ProgStart := TRUE;
   END_IF;
   // 含义：将 (((#HorDrillStep.S12 AND "DB1080_Component".Robot.Status.Busy) AND "DB1081_ValveCall".ST01.Z05.ExtPos) AND "DB1900_Communication_PC".Para.ProduceMode2) OR ((((#HorDrillStep.S12 AND "DB1080_Component".Robot.Status.Busy) AND "DB1081_ValveCall".ST01.Z05.ExtPos) AND "DB1900_Communication_PC".Para.ProduceMode3) AND "DB720_KuKa_MainCtrl".StatusIn.do_Gouge_Pos) OR ((((#HorDrillStep.S12 AND "DB1080_Component".Robot.Status.Busy) AND "DB1081_ValveCall".ST01.Z05.ExtPos) AND "DB1900_Communication_PC".Para.ProduceMode3) AND "DB2500 Visual Chiseling".VisualChiselingMode) OR (#HorDrillStep.S12 AND #HorDrillStep.S15) 赋给 #HorDrillStep.S15
   #HorDrillStep.S15 := (((#HorDrillStep.S12 AND "DB1080_Component".Robot.Status.Busy) AND "DB1081_ValveCall".ST01.Z05.ExtPos) AND "DB1900_Communication_PC".Para.ProduceMode2) OR ((((#HorDrillStep.S12 AND "DB1080_Component".Robot.Status.Busy) AND "DB1081_ValveCall".ST01.Z05.ExtPos) AND "DB1900_Communication_PC".Para.ProduceMode3) AND "DB720_KuKa_MainCtrl".StatusIn.do_Gouge_Pos) OR ((((#HorDrillStep.S12 AND "DB1080_Component".Robot.Status.Busy) AND "DB1081_ValveCall".ST01.Z05.ExtPos) AND "DB1900_Communication_PC".Para.ProduceMode3) AND "DB2500 Visual Chiseling".VisualChiselingMode) OR (#HorDrillStep.S12 AND #HorDrillStep.S15);

   // ---------- 网络 14 ----------
   // 标题：**********************打孔坐标计算************************
   // 注释：水平凿击不计算打孔坐标
   // Core Diamond Drill
   // 32mm: Hor; Heligt:  32.5mm; Length: 50mm 100mm   150mm 250mm
   // 52mm:Down;  Heligt:  65mm; Length: 66.66mm 132.33mmmm   233.67mm
   // 82mm Hor; Height:100mm; Length:100mm 300mm
   // 102mm Hor; Height:80mm; Length:400mm
   // 132mm Hor; Height:125mm; Length:400mm
   // 含义：条件 ((((#HorDrillStep.S15 AND "DB720_KuKa_MainCtrl".StatusIn.do_HorDril_Pos) OR (#HorDrillStep.S15 AND "DB720_KuKa_MainCtrl".StatusIn.do_Gouge_Pos)) AND NOT (#HorDrillStep.S17)) AND ("DB1910_DrillData".HorDrill.PosNo = 0)) 成立时，将 "DB1910_DrillData".HorDrill.CurrentDrillLength 传送到 "DB1910_DrillData".HorDrill.AlreadyDrillLength
   IF ((((#HorDrillStep.S15 AND "DB720_KuKa_MainCtrl".StatusIn.do_HorDril_Pos) OR (#HorDrillStep.S15 AND "DB720_KuKa_MainCtrl".StatusIn.do_Gouge_Pos)) AND NOT (#HorDrillStep.S17)) AND ("DB1910_DrillData".HorDrill.PosNo = 0)) THEN
       "DB1910_DrillData".HorDrill.AlreadyDrillLength := "DB1910_DrillData".HorDrill.CurrentDrillLength;
   END_IF;
   // 含义：条件 ((((#HorDrillStep.S15 AND "DB720_KuKa_MainCtrl".StatusIn.do_HorDril_Pos) OR (#HorDrillStep.S15 AND "DB720_KuKa_MainCtrl".StatusIn.do_Gouge_Pos)) AND NOT (#HorDrillStep.S17)) AND ("DB1910_DrillData".HorDrill.PosNo >= 1)) 成立时，将 ("DB1910_DrillData".HorDrill.AlreadyDrillLength + "DB1910_DrillData".HorDrill.CurrentDrillLength) 传送到 "DB1910_DrillData".HorDrill.AlreadyDrillLength
   IF ((((#HorDrillStep.S15 AND "DB720_KuKa_MainCtrl".StatusIn.do_HorDril_Pos) OR (#HorDrillStep.S15 AND "DB720_KuKa_MainCtrl".StatusIn.do_Gouge_Pos)) AND NOT (#HorDrillStep.S17)) AND ("DB1910_DrillData".HorDrill.PosNo >= 1)) THEN
       "DB1910_DrillData".HorDrill.AlreadyDrillLength := ("DB1910_DrillData".HorDrill.AlreadyDrillLength + "DB1910_DrillData".HorDrill.CurrentDrillLength);
   END_IF;
   // 含义：条件 ((#HorDrillStep.S15 AND "DB720_KuKa_MainCtrl".StatusIn.do_HorDril_Pos) OR (#HorDrillStep.S15 AND "DB720_KuKa_MainCtrl".StatusIn.do_Gouge_Pos)) AND NOT (#HorDrillStep.S17) 成立时，将 ("DB1910_DrillData".HorDrill.PosNo + 1) 传送到 "DB1910_DrillData".HorDrill.PosNo
   IF ((#HorDrillStep.S15 AND "DB720_KuKa_MainCtrl".StatusIn.do_HorDril_Pos) OR (#HorDrillStep.S15 AND "DB720_KuKa_MainCtrl".StatusIn.do_Gouge_Pos)) AND NOT (#HorDrillStep.S17) THEN
       "DB1910_DrillData".HorDrill.PosNo := ("DB1910_DrillData".HorDrill.PosNo + 1);
   END_IF;
   // 含义：将 (#HorDrillStep.S15 AND "DB720_KuKa_MainCtrl".StatusIn.do_HorDril_Pos) OR (#HorDrillStep.S15 AND "DB720_KuKa_MainCtrl".StatusIn.do_Gouge_Pos) 赋给 #HorDrillStep.S17
   #HorDrillStep.S17 := (#HorDrillStep.S15 AND "DB720_KuKa_MainCtrl".StatusIn.do_HorDril_Pos) OR (#HorDrillStep.S15 AND "DB720_KuKa_MainCtrl".StatusIn.do_Gouge_Pos);

   // ---------- 网络 15 ----------
   // 标题：速度分时
   // 含义：本网络为 StructuredText（SCL）原文重建，非 LAD 折叠
   IF #Aux.StartDrill AND
       NOT #HorDrillStep.S22 AND
       NOT "DB720_KuKa_MainCtrl".StatusIn.do_ReqStopDril AND
       "DB720_KuKa_MainCtrl".StatusIn.do_ReqDrilling
   THEN
       #Aux.RobotSpeed := REAL_TO_DINT("DB1080_Component".ClinyderPos.Ctrl_Out.Cur_Val_Out * (-1.0) + 100);
       IF NOT "DB1900_Communication_PC".Para.ProduceMode3 THEN
           IF #Aux.RobotSpeed > 0 THEN
               "DB1080_Component".Robot.CTRL_IN.RobotSpeed := DINT_TO_BYTE((#Aux.RobotSpeed) * "DB1900_Communication_PC".Para.RobotSpeed / 100);
           ELSE
               "DB1080_Component".Robot.CTRL_IN.RobotSpeed := 5;
           END_IF;
       ELSE
           IF #Aux.RobotSpeed > 10 THEN
               "DB1080_Component".Robot.CTRL_IN.RobotSpeed := DINT_TO_BYTE((#Aux.RobotSpeed) * "DB1900_Communication_PC".Para.RobotSpeed / 100);
           ELSE
               "DB1080_Component".Robot.CTRL_IN.RobotSpeed := 20;
           END_IF;
       END_IF;
       IF "DB720_KuKa_MainCtrl".CmdOut.gi_ToolTypeNo = 18 THEN
           IF "DB1080_Component".ClinyderPos.Ctrl_Out.Cur_Val_Out < 30 AND "DB1080_Component".ClinyderPos.Ctrl_Out.Cur_Val_Out >= 15 THEN
               "DB1080_Component".Robot.CTRL_IN.RobotSpeed := 1;
           END_IF;
           IF "DB1080_Component".ClinyderPos.Ctrl_Out.Cur_Val_Out >= 30 THEN
               "DB1080_Component".Robot.CTRL_IN.RobotSpeed := 1;
           END_IF;
       END_IF;
   END_IF;
   IF #HorDrillStep.S12 AND NOT #HorDrillStep.S22 AND "DB1900_Communication_PC".Para.ProduceMode3
       AND "DB720_KuKa_MainCtrl".StatusIn.do_DrillReady_Act AND "DB720_KuKa_MainCtrl".CmdOut.di_ChiselCylinderRet THEN
       "DB1080_Component".Robot.CTRL_IN.RobotSpeed := DINT_TO_BYTE(("DB1900_Communication_PC".Para.RobotSpeed) * 100 / 100);
   END_IF;
   IF "DB720_KuKa_MainCtrl".StatusIn.do_HorDril_Pos THEN
       IF "DB1900_Communication_PC".Para.CurrentMaxLimit > 5.0 THEN
           IF "DB1900_Communication_PC".Recv.Current_2 > ("DB1900_Communication_PC".Para.CurrentMaxLimit - 1.5) THEN
               "DB1080_Component".Robot.CTRL_IN.RobotSpeed := 5;
           END_IF;
       ELSE
           IF "DB1900_Communication_PC".Recv.Current_2 > ("DB1900_Communication_PC".Para.CurrentMaxLimit - 0.5) THEN
               "DB1080_Component".Robot.CTRL_IN.RobotSpeed := 5;
           END_IF;
       END_IF;
   END_IF;

   // ---------- 网络 16 ----------
   // 标题：开始钻孔
   // 含义：将 (#HorDrillStep.S15 AND NOT (#HorDrillStep.S22)) AND NOT ("DB1900_Communication_PC".Para.ProduceMode3) 赋给 "DB720_KuKa_MainCtrl".CmdOut.di_HorDril_Ack
   "DB720_KuKa_MainCtrl".CmdOut.di_HorDril_Ack := (#HorDrillStep.S15 AND NOT (#HorDrillStep.S22)) AND NOT ("DB1900_Communication_PC".Para.ProduceMode3);
   // 含义：将 (#HorDrillStep.S15 AND NOT (#HorDrillStep.S22)) AND "DB1900_Communication_PC".Para.ProduceMode3 赋给 "DB720_KuKa_MainCtrl".CmdOut.di_Gouge_Ack
   "DB720_KuKa_MainCtrl".CmdOut.di_Gouge_Ack := (#HorDrillStep.S15 AND NOT (#HorDrillStep.S22)) AND "DB1900_Communication_PC".Para.ProduceMode3;
   // 含义：将 ((((#HorDrillStep.S15 AND "DB720_KuKa_MainCtrl".StatusIn.do_HorDril_Act) OR (#HorDrillStep.S15 AND "DB1900_Communication_PC".Para.ProduceMode3)) AND NOT ("DB720_KuKa_MainCtrl".StatusIn.do_HorDril_Don)) AND NOT ("DB720_KuKa_MainCtrl".StatusIn.do_Gouge_Don)) OR (#HorDrillStep.S15 AND #HorDrillStep.S20) 赋给 #HorDrillStep.S20
   #HorDrillStep.S20 := ((((#HorDrillStep.S15 AND "DB720_KuKa_MainCtrl".StatusIn.do_HorDril_Act) OR (#HorDrillStep.S15 AND "DB1900_Communication_PC".Para.ProduceMode3)) AND NOT ("DB720_KuKa_MainCtrl".StatusIn.do_HorDril_Don)) AND NOT ("DB720_KuKa_MainCtrl".StatusIn.do_Gouge_Don)) OR (#HorDrillStep.S15 AND #HorDrillStep.S20);

   // ---------- 网络 17 ----------
   // 标题：水平    停止钻孔确认    后开始退枪    直到结束
   // 注释：New Added HDrillEndTime.Q and DB1900.DBX131.1 DrillEndMode in ProduceMode3 by WXY 20220413
   // 含义：条件 ((((((#HorDrillStep.S20 AND NOT (#HorDrillStep.S22)) AND "DB720_KuKa_MainCtrl".StatusIn.do_ReqStopDril) AND NOT ("DB1900_Communication_PC".Para.ProduceMode3)) AND ("DB1900_Communication_PC".Send.ScrLen >= #Aux.DrillDepthMin))) AND NOT ("DB1900_Communication_PC".Para.DrillEndMode)) OR (((((#HorDrillStep.S20 AND NOT (#HorDrillStep.S22)) AND "DB720_KuKa_MainCtrl".StatusIn.do_ReqStopDril) AND NOT ("DB1900_Communication_PC".Para.ProduceMode3)) AND "DB1042_Timer".HDrillEndTime.Q) AND "DB1900_Communication_PC".Para.DrillEndMode) OR (((((#HorDrillStep.S20 AND NOT (#HorDrillStep.S22)) AND "DB720_KuKa_MainCtrl".StatusIn.do_ReqStopDril) AND "DB1900_Communication_PC".Para.ProduceMode3) AND "DB1042_Timer".HDrillEndTime.Q) AND "DB1900_Communication_PC".Para.DrillEndMode) OR (((((#HorDrillStep.S20 AND NOT (#HorDrillStep.S22)) AND "DB720_KuKa_MainCtrl".StatusIn.do_ReqStopDril) AND "DB1900_Communication_PC".Para.ProduceMode3) AND ("DB1900_Communication_PC".Send.ScrLen >= "DB1900_Communication_PC".Para.DrillDepth))) OR ((#HorDrillStep.S20 AND NOT (#HorDrillStep.S22)) AND #HorDrillStep.StopDrill_End) OR ((#HorDrillStep.S20 AND NOT (#HorDrillStep.S22)) AND #HorDrillStep.GougeStopDrill_End) 成立时，将 TRUE 传送到 #HorDrillStep.StopDrill_Ack
   IF ((((((#HorDrillStep.S20 AND NOT (#HorDrillStep.S22)) AND "DB720_KuKa_MainCtrl".StatusIn.do_ReqStopDril) AND NOT ("DB1900_Communication_PC".Para.ProduceMode3)) AND ("DB1900_Communication_PC".Send.ScrLen >= #Aux.DrillDepthMin))) AND NOT ("DB1900_Communication_PC".Para.DrillEndMode)) OR (((((#HorDrillStep.S20 AND NOT (#HorDrillStep.S22)) AND "DB720_KuKa_MainCtrl".StatusIn.do_ReqStopDril) AND NOT ("DB1900_Communication_PC".Para.ProduceMode3)) AND "DB1042_Timer".HDrillEndTime.Q) AND "DB1900_Communication_PC".Para.DrillEndMode) OR (((((#HorDrillStep.S20 AND NOT (#HorDrillStep.S22)) AND "DB720_KuKa_MainCtrl".StatusIn.do_ReqStopDril) AND "DB1900_Communication_PC".Para.ProduceMode3) AND "DB1042_Timer".HDrillEndTime.Q) AND "DB1900_Communication_PC".Para.DrillEndMode) OR (((((#HorDrillStep.S20 AND NOT (#HorDrillStep.S22)) AND "DB720_KuKa_MainCtrl".StatusIn.do_ReqStopDril) AND "DB1900_Communication_PC".Para.ProduceMode3) AND ("DB1900_Communication_PC".Send.ScrLen >= "DB1900_Communication_PC".Para.DrillDepth))) OR ((#HorDrillStep.S20 AND NOT (#HorDrillStep.S22)) AND #HorDrillStep.StopDrill_End) OR ((#HorDrillStep.S20 AND NOT (#HorDrillStep.S22)) AND #HorDrillStep.GougeStopDrill_End) THEN
       #HorDrillStep.StopDrill_Ack := TRUE;
   END_IF;
   // 含义：将 ((#HorDrillStep.S20 AND NOT ("DB1900_Communication_PC".Para.ProduceMode3)) AND "DB720_KuKa_MainCtrl".StatusIn.do_HorDril_Don) OR ((#HorDrillStep.S20 AND "DB1900_Communication_PC".Para.ProduceMode3) AND "DB720_KuKa_MainCtrl".StatusIn.do_Gouge_Don) OR ((#HorDrillStep.S20 AND "DB1900_Communication_PC".Para.ProduceMode3) AND "DB720_KuKa_MainCtrl".StatusIn.do_Gouge_Don1) OR (#HorDrillStep.S20 AND "DB1042_Timer".HorChiselTimeOut.Q) OR (#HorDrillStep.S20 AND #HorDrillStep.S22) 赋给 #HorDrillStep.S22
   #HorDrillStep.S22 := ((#HorDrillStep.S20 AND NOT ("DB1900_Communication_PC".Para.ProduceMode3)) AND "DB720_KuKa_MainCtrl".StatusIn.do_HorDril_Don) OR ((#HorDrillStep.S20 AND "DB1900_Communication_PC".Para.ProduceMode3) AND "DB720_KuKa_MainCtrl".StatusIn.do_Gouge_Don) OR ((#HorDrillStep.S20 AND "DB1900_Communication_PC".Para.ProduceMode3) AND "DB720_KuKa_MainCtrl".StatusIn.do_Gouge_Don1) OR (#HorDrillStep.S20 AND "DB1042_Timer".HorChiselTimeOut.Q) OR (#HorDrillStep.S20 AND #HorDrillStep.S22);
   // 含义：条件 ((#HorDrillStep.S20 AND NOT ("DB1900_Communication_PC".Para.ProduceMode3)) AND "DB720_KuKa_MainCtrl".StatusIn.do_HorDril_Don) OR ((#HorDrillStep.S20 AND "DB1900_Communication_PC".Para.ProduceMode3) AND "DB720_KuKa_MainCtrl".StatusIn.do_Gouge_Don) OR ((#HorDrillStep.S20 AND "DB1900_Communication_PC".Para.ProduceMode3) AND "DB720_KuKa_MainCtrl".StatusIn.do_Gouge_Don1) OR (#HorDrillStep.S20 AND "DB1042_Timer".HorChiselTimeOut.Q) OR (#HorDrillStep.S20 AND #HorDrillStep.S22) 成立时，将 FALSE 传送到 #HorDrillStep.StopDrill_Ack
   IF ((#HorDrillStep.S20 AND NOT ("DB1900_Communication_PC".Para.ProduceMode3)) AND "DB720_KuKa_MainCtrl".StatusIn.do_HorDril_Don) OR ((#HorDrillStep.S20 AND "DB1900_Communication_PC".Para.ProduceMode3) AND "DB720_KuKa_MainCtrl".StatusIn.do_Gouge_Don) OR ((#HorDrillStep.S20 AND "DB1900_Communication_PC".Para.ProduceMode3) AND "DB720_KuKa_MainCtrl".StatusIn.do_Gouge_Don1) OR (#HorDrillStep.S20 AND "DB1042_Timer".HorChiselTimeOut.Q) OR (#HorDrillStep.S20 AND #HorDrillStep.S22) THEN
       #HorDrillStep.StopDrill_Ack := FALSE;
   END_IF;

   // ---------- 网络 18 ----------
   // 标题：斜打    停止钻孔确认    后开始退枪    直到结束
   // 注释：Recv.Current DB1900.DBD116 <  CurrentMinLimit DB1900.DBD218  cgange to Recv.Current DB1900.DBD116 <  CurrentMinLimit DB1900.DBD218  by WXY 20220413
   // 含义：将 (((((#HorDrillStep.S22 AND NOT (#HorDrillStep.S25)) AND "DB1900_Communication_PC".Para.ProduceMode3) AND "DB720_KuKa_MainCtrl".StatusIn.do_ReqStopDril) AND ("DB1900_Communication_PC".Send.ScrLen >= #Aux.DrillDepthMin))) OR ((((#HorDrillStep.S22 AND NOT (#HorDrillStep.S25)) AND "DB1900_Communication_PC".Para.ProduceMode3) AND "DB720_KuKa_MainCtrl".StatusIn.do_ReqStopDril) AND "DB1042_Timer".GougeTimeOut_1.Q) OR ((((#HorDrillStep.S22 AND NOT (#HorDrillStep.S25)) AND "DB1900_Communication_PC".Para.ProduceMode3) AND "DB720_KuKa_MainCtrl".StatusIn.do_ReqStopDril) AND "DB1042_Timer".GougeTimeOut_2.Q) OR ((((#HorDrillStep.S22 AND NOT (#HorDrillStep.S25)) AND "DB1900_Communication_PC".Para.ProduceMode3) AND "DB720_KuKa_MainCtrl".StatusIn.do_ReqStopDril) AND #HorDrillStep.GougeStopDrill_End) 赋给 #HorDrillStep.GougeStopDrill_Ack
   #HorDrillStep.GougeStopDrill_Ack := (((((#HorDrillStep.S22 AND NOT (#HorDrillStep.S25)) AND "DB1900_Communication_PC".Para.ProduceMode3) AND "DB720_KuKa_MainCtrl".StatusIn.do_ReqStopDril) AND ("DB1900_Communication_PC".Send.ScrLen >= #Aux.DrillDepthMin))) OR ((((#HorDrillStep.S22 AND NOT (#HorDrillStep.S25)) AND "DB1900_Communication_PC".Para.ProduceMode3) AND "DB720_KuKa_MainCtrl".StatusIn.do_ReqStopDril) AND "DB1042_Timer".GougeTimeOut_1.Q) OR ((((#HorDrillStep.S22 AND NOT (#HorDrillStep.S25)) AND "DB1900_Communication_PC".Para.ProduceMode3) AND "DB720_KuKa_MainCtrl".StatusIn.do_ReqStopDril) AND "DB1042_Timer".GougeTimeOut_2.Q) OR ((((#HorDrillStep.S22 AND NOT (#HorDrillStep.S25)) AND "DB1900_Communication_PC".Para.ProduceMode3) AND "DB720_KuKa_MainCtrl".StatusIn.do_ReqStopDril) AND #HorDrillStep.GougeStopDrill_End);
   // 含义：调用计数器实例 "DB1042_Timer".GougeTimeOut_1.TON（上升沿计数，当前值写入 CV）
   "DB1042_Timer".GougeTimeOut_1.TON(IN := ((((#HorDrillStep.S22 AND NOT (#HorDrillStep.S25)) AND "DB1900_Communication_PC".Para.ProduceMode3) AND "DB720_KuKa_MainCtrl".StatusIn.do_ReqStopDril) AND ("DB1900_Communication_PC".Recv.Current_2 > "DB1900_Communication_PC".Para.CurrentMinLimit)),
                                     PT := T#3S);
   // 含义：调用定时器实例 "DB1042_Timer".GougeTimeOut_2.TON
   "DB1042_Timer".GougeTimeOut_2.TON(IN := ((#HorDrillStep.S22 AND NOT (#HorDrillStep.S25)) AND "DB1900_Communication_PC".Para.ProduceMode3) AND "DB720_KuKa_MainCtrl".StatusIn.do_ReqStopDril,
                                     PT := T#6S);
   // 含义：将 ((#HorDrillStep.S22 AND "DB1900_Communication_PC".Para.ProduceMode3) AND "DB720_KuKa_MainCtrl".StatusIn.do_Gouge_Don1) OR (#HorDrillStep.S22 AND NOT ("DB1900_Communication_PC".Para.ProduceMode3)) OR (#HorDrillStep.S22 AND #HorDrillStep.S25) 赋给 #HorDrillStep.S25
   #HorDrillStep.S25 := ((#HorDrillStep.S22 AND "DB1900_Communication_PC".Para.ProduceMode3) AND "DB720_KuKa_MainCtrl".StatusIn.do_Gouge_Don1) OR (#HorDrillStep.S22 AND NOT ("DB1900_Communication_PC".Para.ProduceMode3)) OR (#HorDrillStep.S22 AND #HorDrillStep.S25);

   // ---------- 网络 19 ----------
   // 标题：**********************钻孔结束，枪退出速度给定*****************************************
   // 含义：条件 ((((((#HorDrillStep.S20 AND NOT (#HorDrillStep.S22)) AND ("DB720_KuKa_MainCtrl".CmdOut.gi_ToolTypeNo = 2))) AND #HorDrillStep.StopDrill_Ack) AND NOT ("DB1900_Communication_PC".Para.ProduceMode3)) AND ("DB1900_Communication_PC".Para.DrillWidth = 22.0)) 成立时，将 25 传送到 "DB1080_Component".Robot.CTRL_IN.RobotSpeed
   IF ((((((#HorDrillStep.S20 AND NOT (#HorDrillStep.S22)) AND ("DB720_KuKa_MainCtrl".CmdOut.gi_ToolTypeNo = 2))) AND #HorDrillStep.StopDrill_Ack) AND NOT ("DB1900_Communication_PC".Para.ProduceMode3)) AND ("DB1900_Communication_PC".Para.DrillWidth = 22.0)) THEN
       "DB1080_Component".Robot.CTRL_IN.RobotSpeed := 25;
   END_IF;
   // 含义：条件 ((((((#HorDrillStep.S20 AND NOT (#HorDrillStep.S22)) AND ("DB720_KuKa_MainCtrl".CmdOut.gi_ToolTypeNo = 2))) AND #HorDrillStep.StopDrill_Ack) AND NOT ("DB1900_Communication_PC".Para.ProduceMode3)) AND ("DB1900_Communication_PC".Para.DrillWidth = 25.0)) 成立时，将 30 传送到 "DB1080_Component".Robot.CTRL_IN.RobotSpeed
   IF ((((((#HorDrillStep.S20 AND NOT (#HorDrillStep.S22)) AND ("DB720_KuKa_MainCtrl".CmdOut.gi_ToolTypeNo = 2))) AND #HorDrillStep.StopDrill_Ack) AND NOT ("DB1900_Communication_PC".Para.ProduceMode3)) AND ("DB1900_Communication_PC".Para.DrillWidth = 25.0)) THEN
       "DB1080_Component".Robot.CTRL_IN.RobotSpeed := 30;
   END_IF;
   // 含义：条件 ((((((#HorDrillStep.S20 AND NOT (#HorDrillStep.S22)) AND ("DB720_KuKa_MainCtrl".CmdOut.gi_ToolTypeNo = 2))) AND #HorDrillStep.StopDrill_Ack) AND NOT ("DB1900_Communication_PC".Para.ProduceMode3)) AND ("DB1900_Communication_PC".Para.DrillWidth > 25.0)) 成立时，将 40 传送到 "DB1080_Component".Robot.CTRL_IN.RobotSpeed
   IF ((((((#HorDrillStep.S20 AND NOT (#HorDrillStep.S22)) AND ("DB720_KuKa_MainCtrl".CmdOut.gi_ToolTypeNo = 2))) AND #HorDrillStep.StopDrill_Ack) AND NOT ("DB1900_Communication_PC".Para.ProduceMode3)) AND ("DB1900_Communication_PC".Para.DrillWidth > 25.0)) THEN
       "DB1080_Component".Robot.CTRL_IN.RobotSpeed := 40;
   END_IF;
   // 含义：条件 (((((#HorDrillStep.S20 AND NOT (#HorDrillStep.S22)) AND ("DB720_KuKa_MainCtrl".CmdOut.gi_ToolTypeNo = 2))) AND #HorDrillStep.StopDrill_Ack) AND "DB1900_Communication_PC".Para.ProduceMode3) AND "DB1900_Communication_PC".Para.SwingOn 成立时，将 "DB1900_Communication_PC".Para.SwingSpeed 传送到 "DB1080_Component".Robot.CTRL_IN.RobotSpeed
   IF (((((#HorDrillStep.S20 AND NOT (#HorDrillStep.S22)) AND ("DB720_KuKa_MainCtrl".CmdOut.gi_ToolTypeNo = 2))) AND #HorDrillStep.StopDrill_Ack) AND "DB1900_Communication_PC".Para.ProduceMode3) AND "DB1900_Communication_PC".Para.SwingOn THEN
       "DB1080_Component".Robot.CTRL_IN.RobotSpeed := "DB1900_Communication_PC".Para.SwingSpeed;
   END_IF;
   // 含义：条件 (((((#HorDrillStep.S20 AND NOT (#HorDrillStep.S22)) AND ("DB720_KuKa_MainCtrl".CmdOut.gi_ToolTypeNo = 2))) AND #HorDrillStep.StopDrill_Ack) AND "DB1900_Communication_PC".Para.ProduceMode3) AND NOT ("DB1900_Communication_PC".Para.SwingOn) 成立时，将 50 传送到 "DB1080_Component".Robot.CTRL_IN.RobotSpeed
   IF (((((#HorDrillStep.S20 AND NOT (#HorDrillStep.S22)) AND ("DB720_KuKa_MainCtrl".CmdOut.gi_ToolTypeNo = 2))) AND #HorDrillStep.StopDrill_Ack) AND "DB1900_Communication_PC".Para.ProduceMode3) AND NOT ("DB1900_Communication_PC".Para.SwingOn) THEN
       "DB1080_Component".Robot.CTRL_IN.RobotSpeed := 50;
   END_IF;
   // 含义：条件 ((((((#HorDrillStep.S20 AND NOT (#HorDrillStep.S22)) AND ("DB720_KuKa_MainCtrl".CmdOut.gi_ToolTypeNo = 13))) AND #Aux.StartDrill) AND NOT (#HorDrillStep.StopDrill_Ack)) AND ("DB1900_Communication_PC".Recv.Current_2 > 12.0)) 成立时，将 1 传送到 "DB1080_Component".Robot.CTRL_IN.RobotSpeed
   IF ((((((#HorDrillStep.S20 AND NOT (#HorDrillStep.S22)) AND ("DB720_KuKa_MainCtrl".CmdOut.gi_ToolTypeNo = 13))) AND #Aux.StartDrill) AND NOT (#HorDrillStep.StopDrill_Ack)) AND ("DB1900_Communication_PC".Recv.Current_2 > 12.0)) THEN
       "DB1080_Component".Robot.CTRL_IN.RobotSpeed := 1;
   END_IF;
   // 含义：条件 ((((((#HorDrillStep.S20 AND NOT (#HorDrillStep.S22)) AND ("DB720_KuKa_MainCtrl".CmdOut.gi_ToolTypeNo = 13))) AND #Aux.StartDrill) AND #HorDrillStep.StopDrill_Ack) AND ("DB1900_Communication_PC".Recv.Current_2 < 12.0)) 成立时，将 30 传送到 "DB1080_Component".Robot.CTRL_IN.RobotSpeed
   IF ((((((#HorDrillStep.S20 AND NOT (#HorDrillStep.S22)) AND ("DB720_KuKa_MainCtrl".CmdOut.gi_ToolTypeNo = 13))) AND #Aux.StartDrill) AND #HorDrillStep.StopDrill_Ack) AND ("DB1900_Communication_PC".Recv.Current_2 < 12.0)) THEN
       "DB1080_Component".Robot.CTRL_IN.RobotSpeed := 30;
   END_IF;
   // 含义：条件 ((((((#HorDrillStep.S20 AND NOT (#HorDrillStep.S22)) AND ("DB720_KuKa_MainCtrl".CmdOut.gi_ToolTypeNo = 13))) AND #Aux.StartDrill) AND #HorDrillStep.StopDrill_Ack) AND ("DB1900_Communication_PC".Recv.Current_2 >= 12.0)) 成立时，将 10 传送到 "DB1080_Component".Robot.CTRL_IN.RobotSpeed
   IF ((((((#HorDrillStep.S20 AND NOT (#HorDrillStep.S22)) AND ("DB720_KuKa_MainCtrl".CmdOut.gi_ToolTypeNo = 13))) AND #Aux.StartDrill) AND #HorDrillStep.StopDrill_Ack) AND ("DB1900_Communication_PC".Recv.Current_2 >= 12.0)) THEN
       "DB1080_Component".Robot.CTRL_IN.RobotSpeed := 10;
   END_IF;
   // 含义：条件 (((((#HorDrillStep.S20 AND NOT (#HorDrillStep.S22)) AND ("DB720_KuKa_MainCtrl".CmdOut.gi_ToolTypeNo = 18))) AND #HorDrillStep.StopDrill_Ack) AND ("DB1900_Communication_PC".Para.DrillDepth < 100.0)) 成立时，将 20 传送到 "DB1080_Component".Robot.CTRL_IN.RobotSpeed
   IF (((((#HorDrillStep.S20 AND NOT (#HorDrillStep.S22)) AND ("DB720_KuKa_MainCtrl".CmdOut.gi_ToolTypeNo = 18))) AND #HorDrillStep.StopDrill_Ack) AND ("DB1900_Communication_PC".Para.DrillDepth < 100.0)) THEN
       "DB1080_Component".Robot.CTRL_IN.RobotSpeed := 20;
   END_IF;
   // 含义：条件 (((((#HorDrillStep.S20 AND NOT (#HorDrillStep.S22)) AND ("DB720_KuKa_MainCtrl".CmdOut.gi_ToolTypeNo = 18))) AND #HorDrillStep.StopDrill_Ack) AND ("DB1900_Communication_PC".Para.DrillDepth >= 100.0)) 成立时，将 30 传送到 "DB1080_Component".Robot.CTRL_IN.RobotSpeed
   IF (((((#HorDrillStep.S20 AND NOT (#HorDrillStep.S22)) AND ("DB720_KuKa_MainCtrl".CmdOut.gi_ToolTypeNo = 18))) AND #HorDrillStep.StopDrill_Ack) AND ("DB1900_Communication_PC".Para.DrillDepth >= 100.0)) THEN
       "DB1080_Component".Robot.CTRL_IN.RobotSpeed := 30;
   END_IF;

